// TIA Portal V21 export
// export: Created 2000-01-01T00:00:00.0000000Z, ExportSetting None
TYPE "UDT_HMI_RingFifo"
   STRUCT
      bManualEnqueue { ExternalWritable := 'False'} : Bool;   // HMI手动入队触发
      bManualDequeue { ExternalWritable := 'False'} : Bool;   // HMI手动出队触发
      bClearCmd { ExternalWritable := 'False'} : Bool;   // HMI清空队列命令
      diManualItemIn { ExternalWritable := 'False'} : DInt;   // HMI手动入队数值
      diLastItemOut { ExternalWritable := 'False'} : DInt;   // 状态反馈：最近出队数值
      diHeadPreview { ExternalWritable := 'False'} : DInt;   // 状态反馈：队首待出队元素预览
      iCount { ExternalWritable := 'False'} : Int;   // 状态反馈：当前队列元素数量
      bIsEmpty { ExternalWritable := 'False'} : Bool;   // 状态反馈：队列空
      bIsFull { ExternalWritable := 'False'} : Bool;   // 状态反馈：队列满
      bError { ExternalWritable := 'False'} : Bool;   // 状态反馈：溢出或下溢错误
      wStatus { ExternalWritable := 'False'} : Word;   // 状态码：16#0000正常, 16#8001满入溢出, 16#8002空出下溢
   END_STRUCT;
END_TYPE
